// TIA Portal V21 export
// export: Created 2026-08-21T20:18:49.2416972Z, ExportSetting None, DisplayName Totally Integrated Automation Portal, DisplayVersion V21, DisplayName STEP 7 Professional, DisplayVersion V21, DisplayName STEP 7 Safety, DisplayVersion V21, DisplayName Tech WebApplication, DisplayVersion V21, DisplayName WinCC Basic/Comfort/Advanced, DisplayVersion V21, DisplayName WinCC Professional, DisplayVersion V21, DisplayName WinCC Unified, DisplayVersion V21
FUNCTION_BLOCK "PT1"   // FB4, SCL
{ S7_Optimized_Access := 'TRUE' }
// stored: MemoryReserve 100, SetENOAutomatically false
   VAR_INPUT
      On { ExternalAccessible := 'False'; ExternalVisible := 'False'; ExternalWritable := 'False'} : Bool;   // 0 = Off => In = 0.0
      In_Raw { ExternalAccessible := 'False'; ExternalVisible := 'False'; ExternalWritable := 'False'} : Int;
      P { ExternalAccessible := 'False'; ExternalVisible := 'False'; ExternalWritable := 'False'} : Real := 1.0;   // Propotional parameter
      T { ExternalAccessible := 'False'; ExternalVisible := 'False'; ExternalWritable := 'False'} : Real := 1.0;   // Time constant [s]
      t_cyc { ExternalAccessible := 'False'; ExternalVisible := 'False'; ExternalWritable := 'False'} : Real := 0.1;   // OB-Cycle time
   END_VAR
   VAR_OUTPUT
      Out { ExternalAccessible := 'False'; ExternalVisible := 'False'; ExternalWritable := 'False'} : Real := 0.0;
      Out_Raw : Int := 0;
   END_VAR
   VAR
      "Out-1" { ExternalAccessible := 'False'; ExternalVisible := 'False'; ExternalWritable := 'False'} : Real := 0.0;
   END_VAR
BEGIN
   IF #On THEN
       #Out_Raw := #"Out-1" + (#P * (#In_Raw - #"Out-1") * (#t_cyc / (#T + #t_cyc)));
   ELSE
       #Out_Raw := #"Out-1" + (#P * (0.0 - #"Out-1") * (#t_cyc / (#T + #t_cyc)));
   END_IF;

   #"Out-1" := #Out_Raw; //Save output value end of this cycle
   #Out := (INT_TO_REAL(#Out_Raw) / 27648) * 100;
END_FUNCTION_BLOCK
